Fanuc KAREL source: kb00111.compact.KL

PROGRAM KB00111
%STACKSIZE=65535
%PRIORITY=65535
%NOLOCKGROUP
VAR
P1 : FILE
RESULT : INTEGER
BEGIN
RESULT=IO_STATUS(P1)
END KB00111
